{region 'Documentation'}
(*!
<summary>Checks the untouched declaration snapshot through direct and interface reads; never calls the subject.</summary>
*)
{endregion}
FUNCTION_BLOCK Test_PreparationInitialStatus EXTENDS TestCaseBase
VAR
    FSubject : PreparationStatusProbe;
    FView : I_Preparation;
    FSnapshotCopy : ST_PreparationStatus;
    FObserved : ST_PreparationStatus;
    FExpected : ST_PreparationStatus;
    FObservedEnabled : BOOL;
    FExpectedEnabled : BOOL;
    FCheckPerformed : BOOL;
    FObservedCallCount : UDINT;
    FExpectedCallCount : UDINT;
    FCheckDiagnosticState : AssertEqual_Int;
    FCheckExecutionStatus : AssertEqual_Int;
    FCheckReady : AssertEqual_Bool;
    FCheckRunning : AssertEqual_Bool;
    FCheckCompleted : AssertEqual_Bool;
    FCheckError : AssertEqual_Bool;
    FCheckEnabled : AssertEqual_Bool;
    FCheckCallCount : AssertEqual_UDInt;
    FCheckCopyDetached : AssertEqual_Bool;
END_VAR
VAR CONSTANT
    DirectObservation : E_State := E_State.Running;
    DetachedSnapshot : E_State := E_State.Running + 1;
END_VAR

SUPER^();

{region 'Documentation'}
(*!
<summary>Contributes all owned Assertion results without executing the subjects.</summary>
*)
{endregion}
METHOD PROTECTED AggregateResults
VAR_INPUT
    Aggregator : I_ResultAggregator; //! Borrowed result sink owned by the outer Test Case; add this test's checking Assertions without resetting or retaining the sink.
END_VAR
Aggregator.AddProvider(Provider := FCheckDiagnosticState);
Aggregator.AddProvider(Provider := FCheckExecutionStatus);
Aggregator.AddProvider(Provider := FCheckReady);
Aggregator.AddProvider(Provider := FCheckRunning);
Aggregator.AddProvider(Provider := FCheckCompleted);
Aggregator.AddProvider(Provider := FCheckError);
Aggregator.AddProvider(Provider := FCheckEnabled);
Aggregator.AddProvider(Provider := FCheckCallCount);
Aggregator.AddProvider(Provider := FCheckCopyDetached);
END_METHOD

{region 'Documentation'}
(*!
<summary>Requires valid base configuration and every owned Assertion.</summary>
*)
{endregion}
METHOD PROTECTED CheckInitialization : BOOL //! TRUE when the inherited initialization check and this concrete fixture check both accept the setup.
CheckInitialization := FALSE;
IF NOT SUPER^.CheckInitialization() THEN
    RETURN;
END_IF;
IF NOT FCheckDiagnosticState.IsInitialized
    OR NOT FCheckExecutionStatus.IsInitialized
    OR NOT FCheckReady.IsInitialized
    OR NOT FCheckRunning.IsInitialized
    OR NOT FCheckCompleted.IsInitialized
    OR NOT FCheckError.IsInitialized
    OR NOT FCheckEnabled.IsInitialized
    OR NOT FCheckCallCount.IsInitialized
    OR NOT FCheckCopyDetached.IsInitialized THEN
    RETURN;
END_IF;

CheckInitialization := TRUE;
END_METHOD

{region 'Documentation'}
(*!
<summary>Configures this scenario, its local subjects and named Assertions.</summary>
*)
{endregion}
METHOD PROTECTED Configure
FPreparationStateCount := 0;
FTestStateCount := 2;
FCheckPerformed := FALSE;
FView := FSubject;
FSnapshotCopy.Completed := FALSE;

FCheckDiagnosticState.Initialize(Parent := THIS^,
    AssertionName := 'DiagnosticState');
FCheckExecutionStatus.Initialize(Parent := THIS^,
    AssertionName := 'ExecutionStatus');
FCheckReady.Initialize(Parent := THIS^,
    AssertionName := 'Ready');
FCheckRunning.Initialize(Parent := THIS^,
    AssertionName := 'Running');
FCheckCompleted.Initialize(Parent := THIS^,
    AssertionName := 'Completed');
FCheckError.Initialize(Parent := THIS^,
    AssertionName := 'Error');
FCheckEnabled.Initialize(Parent := THIS^,
    AssertionName := 'Enabled');
FCheckCallCount.Initialize(Parent := THIS^,
    AssertionName := 'CallCount');
FCheckCopyDetached.Initialize(Parent := THIS^,
    AssertionName := 'CopyDetached');
END_METHOD

{region 'Documentation'}
(*!
<summary>Ends scenario processing without issuing further resource commands.</summary>
*)
{endregion}
METHOD PROTECTED ProcessAbort
VAR_INPUT
    Enable : BOOL; //! Phase permission supplied by the owning Test Case; FALSE does not authorize progression, while observation may continue.
END_VAR
IF Enable THEN
    CompleteAbort();
END_IF;
END_METHOD

{region 'Documentation'}
(*!
<summary>Compares independent expected values with the captured observations; called when disabled as well.</summary>
*)
{endregion}
METHOD PROTECTED ProcessAssertions
VAR_INPUT
    Enable : BOOL; //! Phase permission supplied by the owning Test Case; FALSE does not authorize progression, while observation may continue.
END_VAR
FCheckDiagnosticState(Enable := Enable,
    State := State,
    IN := TO_INT(FObserved.State),
    Expected := TO_INT(FExpected.State));

FCheckExecutionStatus(Enable := Enable,
    State := State,
    IN := TO_INT(FObserved.ExecutionStatus),
    Expected := TO_INT(FExpected.ExecutionStatus));

FCheckReady(Enable := Enable,
    State := State,
    IN := FObserved.Ready,
    Expected := FExpected.Ready);

FCheckRunning(Enable := Enable,
    State := State,
    IN := FObserved.Running,
    Expected := FExpected.Running);

FCheckCompleted(Enable := Enable,
    State := State,
    IN := FObserved.Completed,
    Expected := FExpected.Completed);

FCheckError(Enable := Enable,
    State := State,
    IN := FObserved.Error,
    Expected := FExpected.Error);

FCheckEnabled(Enable := Enable,
    State := State,
    IN := FObservedEnabled,
    Expected := FExpectedEnabled);

FCheckCallCount(Enable := Enable,
    State := State,
    IN := FObservedCallCount,
    Expected := FExpectedCallCount);

FCheckCopyDetached(Enable := Enable,
    State := State,
    IN := FSnapshotCopy.Completed,
    Expected := State = DetachedSnapshot);

IF Enable
    AND FCheckDiagnosticState.EvaluationActive
    AND FCheckExecutionStatus.EvaluationActive
    AND FCheckReady.EvaluationActive
    AND FCheckRunning.EvaluationActive
    AND FCheckCompleted.EvaluationActive
    AND FCheckError.EvaluationActive
    AND FCheckEnabled.EvaluationActive
    AND FCheckCallCount.EvaluationActive
    AND FCheckCopyDetached.EvaluationActive THEN
    FCheckPerformed := TRUE;
END_IF;
END_METHOD

{region 'Documentation'}
(*!
<summary>Subjects are exercised by the test, not used as its start prerequisite.</summary>
*)
{endregion}
METHOD PROTECTED ProcessPreparations
VAR_INPUT
    // SA0033: Required hook; this scenario has no Preparation phase.
    {attribute 'analysis' := '-33'}
    Enable : BOOL; //! Phase permission supplied by the owning Test Case; FALSE does not authorize progression, while observation may continue.
END_VAR
END_METHOD

{region 'Documentation'}
(*!
<summary>Restores repeatable fixture state and resets Assertions before returning to Idle.</summary>
*)
{endregion}
METHOD PROTECTED ProcessReset
FCheckPerformed := FALSE;
FSnapshotCopy.Completed := FALSE;
FCheckDiagnosticState.Reset();
FCheckExecutionStatus.Reset();
FCheckReady.Reset();
FCheckRunning.Reset();
FCheckCompleted.Reset();
FCheckError.Reset();
FCheckEnabled.Reset();
FCheckCallCount.Reset();
FCheckCopyDetached.Reset();
CompleteReset();
END_METHOD

{region 'Documentation'}
(*!
<summary>Exercises one named scenario step per call; advances only after actual Assertion evaluation.</summary>
*)
{endregion}
METHOD PROTECTED ProcessTests
VAR_INPUT
    Enable : BOOL; //! Phase permission supplied by the owning Test Case; FALSE does not authorize progression, while observation may continue.
END_VAR
IF NOT Enable THEN
    RETURN;
END_IF;

IF FCheckPerformed THEN
    FCheckPerformed := FALSE;
    IF State = DetachedSnapshot THEN
        CompleteTests();
        RETURN;
    END_IF;
    NextTestState();
    IF NOT IsTestingActive THEN
        RETURN;
    END_IF;
END_IF;

CASE State OF
    DirectObservation:
        FObserved := FSubject.Status;
        FObservedEnabled := FSubject.Enabled;
        FExpected.State := E_State.Uninitialized;
        FExpected.ExecutionStatus := E_ExecutionStatus.Unknown;
        FExpected.Ready := FALSE;
        FExpected.Running := FALSE;
        FExpected.Completed := FALSE;
        FExpected.Error := FALSE;
        FExpectedEnabled := FALSE;
        FExpectedCallCount := 0;

    DetachedSnapshot:
        FSnapshotCopy := FView.Status;
        FSnapshotCopy.Completed := TRUE;
        FObserved := FView.Status;
        FObservedEnabled := FSubject.Enabled;
        FExpected.State := E_State.Uninitialized;
        FExpected.ExecutionStatus := E_ExecutionStatus.Unknown;
        FExpected.Ready := FALSE;
        FExpected.Running := FALSE;
        FExpected.Completed := FALSE;
        FExpected.Error := FALSE;
        FExpectedEnabled := FALSE;
        FExpectedCallCount := 0;

ELSE
    Error(Message := 'Unexpected Preparation test state.');
    RETURN;
END_CASE;

FObservedCallCount := FSubject.CallCount;
END_METHOD

END_FUNCTION_BLOCK

(* stored: Version 1.1.0.1
   POU Test_PreparationInitialStatus: Id {bfdefe4e-2de7-43b1-9e5a-7ccde384ee7c}, SpecialFunc None
   Folder Internal: Id {62d877b6-5c34-4c34-8e2a-cdca12c40910}
   Method AggregateResults: Id {32e72a7c-ca17-46c3-b29c-8f3b4cd87d95}
   Method CheckInitialization: Id {4ae9e8a3-00a9-4d68-a51b-04563adfa7e6}
   Method Configure: Id {dd5eaa9c-0b6a-4eb2-9301-9aadb26b8f06}
   Method ProcessAbort: Id {13714c1b-cd09-4758-8d09-8469765a3288}
   Method ProcessAssertions: Id {325498f2-2652-465b-9790-4982a0fca35e}
   Method ProcessPreparations: Id {17b7ca56-4261-4b6e-9b80-52e481c7eb07}
   Method ProcessReset: Id {2bae657d-a5da-4dc0-935e-411e8256b2f7}
   Method ProcessTests: Id {0445d4d3-55d6-4eae-b80a-c49c51362160} *)
